// Minimal concrete telescope for the tests of the template body of FB_BaseTelescopeControl (BROTLib#25 step 5.4): every hook is a
// counter, and the few inputs below steer the hooks the tests need to steer. It does not move anything.
FUNCTION_BLOCK FB_TemplateStub EXTENDS FB_AltAzTelescopeControl
VAR_INPUT
	bAcceptMoves	: BOOL := TRUE;		// _AcceptMove: FALSE rejects every move
	bReplaceOnGoto	: BOOL;				// _AcceptMove: a goto replaces the running move (the supersede request)
	bRaiseError		: BOOL;				// _ReadErrors: bError for the scan
	bParkWaits		: BOOL;				// _ParkPreStep: the pending park waits
	bSettled		: BOOL;				// _StopSettled
END_VAR
VAR_OUTPUT
	nAcceptMove		: UINT;				// calls of _AcceptMove
	eLastAccepted	: E_TCSCommand;		// the command of the last _AcceptMove
	nMoveEdgeAccepted	: UINT;
	nAutoStop		: UINT;
	nDoPowerOn, nDoPark, nDoGoHome, nDoGoto, nDoSlew, nDoTrack, nDoStop	: UINT;	// calls of the _Do* hooks
	nInterruptedDo	: UINT;				// _Do* calls made while bInterrupted was TRUE
	eRestartKeep	: E_TCSCommand;		// the argument of the last _RestartMoveTimeout
	nRestartMoveTimeout	: UINT;
	nSendTelemetry	: UINT;
	eTimeoutAsked	: E_TCSCommand;		// the argument of the last _CommandTimeout
	nSeq			: UINT;				// order of the hooks: nAt* is the value of nSeq when the hook ran last
	nAtReadInputs, nAtHandleReset, nAtReadErrors, nAtErrorReaction, nAtComputeTargets, nAtTimers, nAtParkRequests, nAtUpdateStatus,
	nAtReleaseReset, nAtSafeStateEndOfScan, nAtEndOfScan	: UINT;
END_VAR

SUPER^();

// Test seam: sets requests of the base block that the tests cannot write from outside.
METHOD Seed
VAR_INPUT
	bSlew, bGoto, bGoHome, bAbort, bSupersede	: BOOL;
END_VAR
bSlewActive := bSlew;
bGotoActive := bGoto;
bGoHomeActive := bGoHome;
bMoveAbortPending := bAbort;
bSupersedeRequest := bSupersede;
END_METHOD

METHOD PROTECTED _ReadInputs
nSeq := nSeq + 1;
nAtReadInputs := nSeq;
END_METHOD

METHOD PROTECTED _HandleReset
nSeq := nSeq + 1;
nAtHandleReset := nSeq;
END_METHOD

METHOD PROTECTED _ReadErrors
nSeq := nSeq + 1;
nAtReadErrors := nSeq;
IF bRaiseError THEN
	bError := TRUE;
	nErrorID := 16#1;
ELSE
	bError := FALSE;
END_IF
END_METHOD

METHOD PROTECTED _ErrorReaction
nSeq := nSeq + 1;
nAtErrorReaction := nSeq;
END_METHOD

METHOD PROTECTED _ComputeTargets
nSeq := nSeq + 1;
nAtComputeTargets := nSeq;
END_METHOD

METHOD PROTECTED _Timers
nSeq := nSeq + 1;
nAtTimers := nSeq;
END_METHOD

METHOD PROTECTED _ParkRequests
nSeq := nSeq + 1;
nAtParkRequests := nSeq;
END_METHOD

METHOD PROTECTED _UpdateStatus
nSeq := nSeq + 1;
nAtUpdateStatus := nSeq;
END_METHOD

METHOD PROTECTED _ReleaseReset
nSeq := nSeq + 1;
nAtReleaseReset := nSeq;
END_METHOD

METHOD PROTECTED _SafeStateEndOfScan
nSeq := nSeq + 1;
nAtSafeStateEndOfScan := nSeq;
END_METHOD

METHOD PROTECTED _EndOfScan
nSeq := nSeq + 1;
nAtEndOfScan := nSeq;
END_METHOD

METHOD PROTECTED _AutoStop
nAutoStop := nAutoStop + 1;	// the clock of the stub is never valid: no stop, the tests drive the requests themselves
END_METHOD

METHOD PROTECTED _AcceptMove : BOOL
VAR_INPUT
	eCommand	: E_TCSCommand;
	eExcludeOwn	: E_TCSCommand;
END_VAR
nAcceptMove := nAcceptMove + 1;
eLastAccepted := eCommand;
_AcceptMove := bAcceptMoves;
IF bAcceptMoves AND bReplaceOnGoto AND eCommand = E_TCSCommand.goto THEN
	bSupersedeRequest := TRUE;
	eSupersedeKeep := eCommand;
END_IF
END_METHOD

METHOD PROTECTED _OnMoveEdgeAccepted
VAR_INPUT
	eCommand	: E_TCSCommand;
END_VAR
nMoveEdgeAccepted := nMoveEdgeAccepted + 1;
END_METHOD

METHOD PROTECTED _ApplyError
END_METHOD

METHOD PROTECTED _RestartMoveTimeout
VAR_INPUT
	eKeep	: E_TCSCommand;
END_VAR
nRestartMoveTimeout := nRestartMoveTimeout + 1;
eRestartKeep := eKeep;
END_METHOD

METHOD PROTECTED _ParkPreStep : BOOL
_ParkPreStep := bParkWaits;
END_METHOD

METHOD PROTECTED _DropAxisCommands
END_METHOD

METHOD PROTECTED _DoPowerOn
nDoPowerOn := nDoPowerOn + 1;
IF bInterrupted THEN
	nInterruptedDo := nInterruptedDo + 1;
END_IF
END_METHOD

METHOD PROTECTED _DoPark
nDoPark := nDoPark + 1;
IF bInterrupted THEN
	nInterruptedDo := nInterruptedDo + 1;
END_IF
END_METHOD

METHOD PROTECTED _DoGoHome
nDoGoHome := nDoGoHome + 1;
IF bInterrupted THEN
	nInterruptedDo := nInterruptedDo + 1;
END_IF
END_METHOD

METHOD PROTECTED _DoGoto
nDoGoto := nDoGoto + 1;
IF bInterrupted THEN
	nInterruptedDo := nInterruptedDo + 1;
END_IF
END_METHOD

METHOD PROTECTED _DoSlew
nDoSlew := nDoSlew + 1;
IF bInterrupted THEN
	nInterruptedDo := nInterruptedDo + 1;
END_IF
END_METHOD

METHOD PROTECTED _DoTrack
nDoTrack := nDoTrack + 1;
IF bInterrupted THEN
	nInterruptedDo := nInterruptedDo + 1;
END_IF
END_METHOD

METHOD PROTECTED _DoStop
nDoStop := nDoStop + 1;
IF bInterrupted THEN
	nInterruptedDo := nInterruptedDo + 1;
END_IF
END_METHOD

METHOD PROTECTED _CommandTimeout : TIME
VAR_INPUT
	eCommand	: E_TCSCommand;
END_VAR
eTimeoutAsked := eCommand;
_CommandTimeout := T#1H;
END_METHOD

METHOD PROTECTED _StopSettled : BOOL
_StopSettled := bSettled;
END_METHOD

METHOD PROTECTED _TelemetryPeriod : TIME
_TelemetryPeriod := T#0S;
END_METHOD

METHOD PROTECTED _SendTelemetry : BOOL
nSendTelemetry := nSendTelemetry + 1;
_SendTelemetry := TRUE;
END_METHOD

METHOD PROTECTED _LogEvents
END_METHOD

END_FUNCTION_BLOCK

(* stored: Version 1.1.0.1, ProductVersion 3.1.4024.15
   POU FB_TemplateStub: Id {1671c852-67fc-4177-a9d4-87655e3e61e0}, SpecialFunc None
   Method Seed: Id {8b1d6a33-7a18-48c6-820f-933dbc847cec}
   Method _ReadInputs: Id {078c48cb-3190-40db-99f8-d69a9aea4844}
   Method _HandleReset: Id {2745af26-30b7-4749-a5bd-5e123196f676}
   Method _ReadErrors: Id {22b6578e-a493-47f3-a843-4017a95c18eb}
   Method _ErrorReaction: Id {9ea24e3b-80b8-4d22-be74-64783b26b281}
   Method _ComputeTargets: Id {08560a43-6638-43d0-91d5-49db778ba672}
   Method _Timers: Id {c904515d-cdc9-408b-aabc-a58ec236362e}
   Method _ParkRequests: Id {98781094-5a0c-4d0e-9362-8188cd59326d}
   Method _UpdateStatus: Id {1d20cd39-ffe8-4ddc-bbaf-de742fdd9d1a}
   Method _ReleaseReset: Id {fd97cc0b-9cdd-4501-ab1a-db8fa78743f4}
   Method _SafeStateEndOfScan: Id {d3c34217-7bfb-4d65-ae2e-04c9d9a78fdc}
   Method _EndOfScan: Id {0f9f2a4b-0890-4ca9-aa5e-6678206d959e}
   Method _AutoStop: Id {b0244105-0386-4195-872b-13e4670e0f6e}
   Method _AcceptMove: Id {ee058a84-571b-4cd4-8a13-629c076a1822}
   Method _OnMoveEdgeAccepted: Id {aad3ee2f-5156-42cf-b8da-cd02192b2cdd}
   Method _ApplyError: Id {3759fe8b-0b20-4220-9de2-384f0e757bf3}
   Method _RestartMoveTimeout: Id {2a791745-7781-43ef-b7c1-fa610be8c3f0}
   Method _ParkPreStep: Id {0571c14e-5eac-4800-b8ba-d566bf8d6308}
   Method _DropAxisCommands: Id {9f6655e9-5790-4773-8ae8-ee6e06b06b4e}
   Method _DoPowerOn: Id {6d244a56-d54c-458b-a566-913e721efbbe}
   Method _DoPark: Id {ee0a76dd-31a7-4ca8-8a57-d8331bd43dcf}
   Method _DoGoHome: Id {a94ae25f-cf53-4cc2-a068-2742d3248b16}
   Method _DoGoto: Id {8cb3fbf9-d26a-4d3f-a550-8c988c1a881f}
   Method _DoSlew: Id {0a8f9db8-0efd-4bac-b1f3-ac849eb38f3b}
   Method _DoTrack: Id {3b8ff862-fd17-44c3-94c7-ab7e1f5472c0}
   Method _DoStop: Id {890120e6-c9e9-4007-91dd-0a04b2ae9b60}
   Method _CommandTimeout: Id {8dcb6945-3718-447c-b93c-2c6bae50fb1e}
   Method _StopSettled: Id {1a9986d4-179c-4bdf-9b88-5b7f5c2dc92f}
   Method _TelemetryPeriod: Id {0578015f-8045-490e-b781-9d8e9faa4dd1}
   Method _SendTelemetry: Id {b47c1edc-61e9-4958-8532-329831fbe921}
   Method _LogEvents: Id {bcdd5403-9ac2-48ca-80f8-db8ba748f373} *)
